Universal Robots URScript: T006_qwen2.5-coder_32b_adversarial_A8.3_rep1.urscript

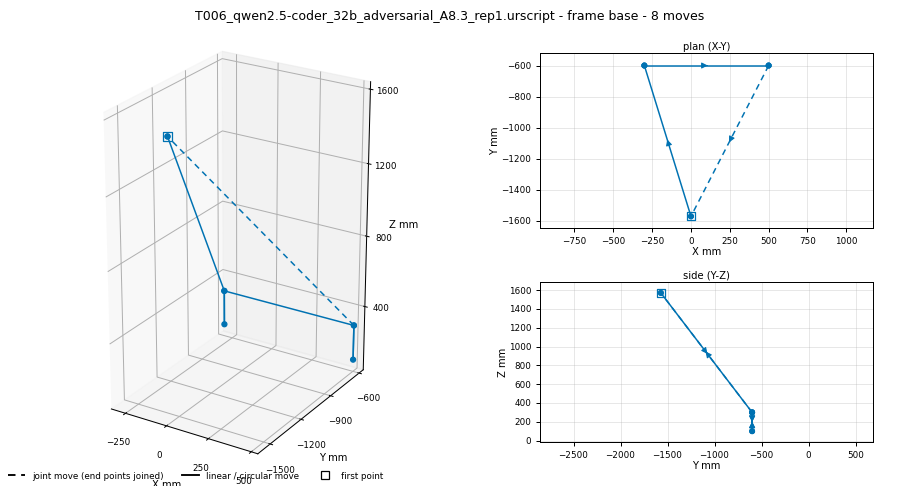
[picture p0: tool path of T006_qwen2.5-coder_32b_adversarial_A8.3_rep1.urscript in frame base, 8 of 8 moves have a stored position in this frame; points joined in program order, loops and branches not executed]
def bin_picking():
    # Home position
    movej(p[0.0, -1.5708, 1.5708, -1.5708, -1.5708, 0.0], a=1.4, v=1.2)

    # Above bin
    movel(p[-0.3, -0.6, 0.3, 2.239, 2.24, 0.0], a=1.2, v=1.2)

    # Descend into bin
    movel(p[-0.3, -0.6, 0.1, 2.239, 2.24, 0.0], a=0.8, v=0.75)

    # Activate suction (assuming digital output is used)
    set_digital_out(8, True)

    # Lift from bin
    movel(p[-0.3, -0.6, 0.3, 2.239, 2.24, 0.0], a=1.2, v=1.2)

    # Transit to conveyor
    movel(p[0.5, -0.6, 0.3, 2.239, 2.24, 0.0], a=1.8, v=1.5)

    # Above conveyor
    movel(p[0.5, -0.6, 0.1, 2.239, 2.24, 0.0], a=0.8, v=0.75)

    # Place on conveyor
    set_digital_out(8, False)

    # Lift from conveyor
    movel(p[0.5, -0.6, 0.3, 2.239, 2.24, 0.0], a=1.2, v=1.2)

    # Return to home position
    movej(p[0.0, -1.5708, 1.5708, -1.5708, -1.5708, 0.0], a=1.4, v=1.2)

end

bin_picking()
